(* IEC 61131-3 sources: sis-interlock-demo/tests/POUs/TruthTables/FB_VoteTable2oo3DADI_Test, 1 file *)

(* ---- Fb2oo3DADIMatchesModel.method.decl.st ---- *)
// AUTO-GENERATED by tools_project/gen_voting_tests.py — не редактировать: правьте генератор или модель
//   tools_project/vote_model.py и запустите python tools_project/gen_voting_tests.py
// FB_Voting, схема 2oo3, политика DA, вход DI: все 512 сочетаний
// (требование × достоверность × запрос байпаса по каналу — для FB_Voting); ожидаемые значения —
// эталонная модель tools_project/vote_model.py. Один AssertEquals_BYTE на строку.
METHOD PRIVATE Fb2oo3DADIMatchesModel
VAR
    fbRig : FB_VoteTableRig;   // стенд таблиц (новый экземпляр на тест)
    bRes  : BYTE;              // код результата строки
END_VAR
